FUNCTION_BLOCK FB_Alarm
VAR_INPUT
	rValue : REAL; // Målt verdi 
	rLimit : REAL; // Maks verdi for BAR og temperatur
	bReset : BOOL; // Denne nulstiller alarmen, denne blir brukt i HMIen
END_VAR
VAR_OUTPUT
	bAlarm  : BOOL;    // TRUE når alarmen er aktiv
END_VAR
VAR
	fbLatch : RS; // Fungerer som minnebryter - Eks: Trykket går under 4 Bar, men alarmen fortsetter å gå, fordi den husker at noe skjedde.
	               // Først når noen trykker reset, slår den seg av.
				   // Det er nettopp det RS gjør. SET slår den på, den blir stående på, og RESET slår den av.
				   // fbLatch er ikke en verdi, men en instans av RS-blokken, altså en egen liten “minnebryter” som lever inne i FB_Alarm
END_VAR

// FB_Alarm er røykvarsleren. Den merker brannen og fortsetter å pipe til noen kvitterer.

//FB_Alarm bestemmer om det er alarm.

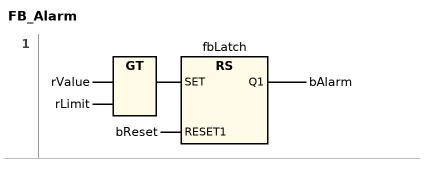
// NETWORK 1
fbLatch(SET := rValue > rLimit, RESET1 := bReset); // RS
bAlarm := fbLatch.Q1;

END_FUNCTION_BLOCK

(* stored: Version 1.1.0.1, ProductVersion 3.1.4026.21
   POU FB_Alarm: Id {e16690ae-fb34-4d5e-8022-4c9ac09ff5f5}, SpecialFunc None *)
